FUNCTION_BLOCK MOD_OccupationIds (* Builds the OPC UA addresses (Occupy, Release, Occupied) and the local channel names of the occupation from the module's name and OPC UA root. Technical: OPC UA and local channel IDs of the occupation *)
  (* Standard: 61499-2 *)
  (* Version 0.1, 2026-09-28, Project contributors, AAU Smart Production Lab *)
  PACKAGE modlib;
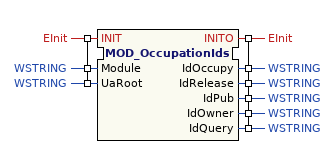
  EVENT_INPUT
    INIT : EInit WITH Module, UaRoot; (* Initialise, once at start-up (the INIT chain); takes the values given with it *)
  END_EVENT
  EVENT_OUTPUT
    INITO : EInit WITH IdOccupy, IdRelease, IdPub, IdOwner, IdQuery; (* Initialised: the next block of the INIT chain goes on *)
  END_EVENT
  VAR_INPUT
    Module : WSTRING; (* The module's name; its local channels are named after it (loc[<Module>/...]) *)
    UaRoot : WSTRING; (* The module's OPC UA folder, e.g. /Objects/Filling *)
  END_VAR
  VAR_OUTPUT
    IdOccupy : WSTRING; (* OPC UA ID of the method Occupy *)
    IdRelease : WSTRING; (* OPC UA ID of the method Release *)
    IdPub : WSTRING; (* OPC UA ID of the published value *)
    IdOwner : WSTRING; (* Local channel of the owner *)
    IdQuery : WSTRING; (* Local channel that asks for the current value (a block that starts later) *)
  END_VAR
  EC_STATES
    INIT : INIT -> INITO;
  END_STATES
  ALGORITHM INIT IN ST:
IdOccupy := CONCAT(CONCAT(CONCAT("opc_ua[CREATE_METHOD;", CONCAT(UaRoot, "/Occupation/")), "Occupy"), "]");
IdRelease := CONCAT(CONCAT(CONCAT("opc_ua[CREATE_METHOD;", CONCAT(UaRoot, "/Occupation/")), "Release"), "]");
IdPub := CONCAT(CONCAT(CONCAT("opc_ua[WRITE;", CONCAT(UaRoot, "/Occupation/")), "Occupied"), "]");
IdOwner := CONCAT(CONCAT("loc[", Module), "/owner]");
IdQuery := CONCAT(CONCAT("loc[", Module), "/owner/query]");
  END_ALGORITHM
END_FUNCTION_BLOCK
